// This function has been automatically generated from the project information.
{attribute 'signature_flag' := '1073741824'}
{attribute 'TcGenerated'}
{attribute 'no-analysis'}
FUNCTION F_GetCompany : WSTRING
VAR_INPUT
	
END_VAR

F_GetCompany := "S&E Engineering";

END_FUNCTION

(* stored: Version 1.1.0.1
   POU F_GetCompany: Id {19107d81-5993-4f52-96a1-49d986f8fbed}, SpecialFunc None *)
